// TIA Portal V21 export
TextList "TL_State"  ListRange=Decimal
  TextListEntry   Text="ISKLJUČENO"
  TextListEntry   From=1, To=1, Text="INICIJALIZACIJA"
  TextListEntry   From=2, To=2, Text="SPREMAN"
  TextListEntry   From=3, To=3, Text="RADI"
  TextListEntry   From=4, To=4, Text="PAUZA"
  TextListEntry   From=5, To=5, Text="ALARM"
  TextListEntry   From=6, To=6, Text="ZAVRŠENO"
  TextListEntry   From=7, To=7, Text="PLANIRANJE"
